(* IEC 61131-3 sources: SemaPLC/sema-plc-benchmark/spec2control-benchmark/data/st-baseline/steel-plant/pous/programs, 9 files *)

(* ---- main.st ---- *)
PROGRAM main
VAR
	Heartbeat : bool;
END_VAR

(* Entry point required by OpenPLC Editor v4. The process sections run as parallel program instances under task0; main only provides a scan heartbeat. *)
Heartbeat := NOT Heartbeat;

END_PROGRAM

(* ---- Section2.st ---- *)
PROGRAM Section2
VAR
	FT101_WildFlow_PV : real;
	FT102_FluxFlow_PV : real;
	TIT101_Temperature_PV : real;
	FFIC103_FluxFlow_SP : real;
	FT_101 : ANALOG_IN;
	FT_102 : ANALOG_IN;
	TIT_101 : ANALOG_IN;
	FFIC_103 : RATIO_CONTROL;
	FIC_102 : PID_BASIC;
	FV_102 : VALVE_ELECTRIC;
	LowFlow_OK_GT : bool;
	FFIC103_LowTempOrLowFlow_OR : bool;
	FFIC103_SensorFaults_OR : bool;
	FFIC103_RangeOrLowTempLowFlow_OR : bool;
	FFIC103_Inhibit_OR : bool;
END_VAR

FT_101(
    PV_Low := 50.0,
    Scaling_Slope := 62.5,
    Scaling_Offset := -250.0,
    Alarm_Enable := TRUE);
FT_102(
    Alarm_Enable := TRUE);
TIT_101(
    PV_Low := 800.0,
    Alarm_Enable := TRUE);
FFIC103_LowTempOrLowFlow_OR := FT_101.Low_Alarm OR TIT_101.Low_Alarm;
FFIC103_RangeOrLowTempLowFlow_OR := FT_101.High_Alarm OR FFIC103_LowTempOrLowFlow_OR;
FFIC103_SensorFaults_OR := FT_101.General_Fault OR FT_102.General_Fault;
FFIC103_Inhibit_OR := FFIC103_SensorFaults_OR OR FFIC103_RangeOrLowTempLowFlow_OR;
LowFlow_OK_GT := (FT_101.PV > 50.0);
FFIC_103(
    Auto := LowFlow_OK_GT,
    PrimaryPV := FT_101.PV,
    SecondaryPV := FT_102.PV,
    RatioSP := 0.4,
    MV_MIN := 200.0,
    MV_MAX := 300.0,
    Inhibit := FFIC103_Inhibit_OR);
FIC_102(
    AUTO := LowFlow_OK_GT,
    PV := FT_102.PV,
    SP := FFIC_103.SlaveSP);
FV_102(
    Control_Signal := FIC_102.XOUT,
    Inhibit := FFIC103_LowTempOrLowFlow_OR);

(* Outputs published to other sections / HMI. *)
FT101_WildFlow_PV := FT_101.PV;
FT102_FluxFlow_PV := FT_102.PV;
TIT101_Temperature_PV := TIT_101.PV;
FFIC103_FluxFlow_SP := FFIC_103.SlaveSP;

END_PROGRAM

(* ---- Section3.st ---- *)
PROGRAM Section3
VAR
	PT_201_VOTE_PV : real;
	TT_201_VOTE_PV : real;
	PT_201A : ANALOG_IN;
	PT_201B : ANALOG_IN;
	PT_201C : ANALOG_IN;
	TT_201A : ANALOG_IN;
	TT_201B : ANALOG_IN;
	TT_201C : ANALOG_IN;
	PT_201_VOTE : VOTING_ANALOG;
	TT_201_VOTE : VOTING_ANALOG;
	P_201 : MOTOR_ON_OFF;
	MO_201 : DIGITAL_IN;
	MO_202 : DIGITAL_IN;
	I_201 : BOOL_INPUT;
	I_202 : BOOL_INPUT;
	SI_201 : BOOL_INPUT;
	SI_202 : BOOL_INPUT;
	PT_GeneralFault : bool;
	MO201_Invert : bool;
	PT_SummaryPre : bool;
	PT_SummaryMasked : bool;
	TT_GeneralFault : bool;
	MO202_Invert : bool;
	TT_SummaryPre : bool;
	TT_SummaryMasked : bool;
	PressureInhibit : bool;
	TemperatureInhibit : bool;
	PumpInhibit : bool;
	PT_PressureHigh : bool;
	TT_TemperatureHigh : bool;
	PT_PressurePermissive : bool;
	TT_TemperaturePermissive : bool;
	StartPermissiveOK : bool;
	StartPermissiveNot : bool;
END_VAR

PT_201A(
    PV_High := 100.0,
    Alarm_Enable := TRUE);
PT_201B(
    PV_High := 100.0,
    Alarm_Enable := TRUE);
PT_201C(
    PV_High := 100.0,
    Alarm_Enable := TRUE);
TT_201A(
    Alarm_Enable := TRUE);
TT_201B(
    Alarm_Enable := TRUE);
TT_201C(
    Alarm_Enable := TRUE);
PT_PressureHigh := (PT_201_VOTE_PV > 100.0);
I_201(
    Bool_In := PT_PressureHigh,
    Alarm_OnTrue := TRUE,
    Latch_Enable := TRUE);
MO_201();
MO201_Invert := NOT MO_201.DI_Out;
PT_GeneralFault := PT_201A.General_Fault OR PT_201B.General_Fault OR PT_201C.General_Fault;
PT_SummaryPre := PT_GeneralFault OR PT_201_VOTE.Alarm_Voting_Error;
PT_SummaryMasked := PT_SummaryPre AND MO201_Invert;
SI_201(
    Bool_In := PT_SummaryMasked,
    Alarm_OnTrue := TRUE,
    Latch_Enable := TRUE);
PressureInhibit := I_201.Bool_Out OR SI_201.Bool_Out;
PT_201_VOTE(
    Input1 := PT_201A.PV,
    Input2 := PT_201B.PV,
    Input3 := PT_201C.PV,
    Deviation_Limit := 5.0,
    Voting_Scheme := '"2oo3"',
    EnableAlarm := TRUE,
    Inhibit := PressureInhibit);
TT_TemperatureHigh := (TT_201_VOTE_PV > 75.0);
I_202(
    Bool_In := TT_TemperatureHigh,
    Alarm_OnTrue := TRUE,
    Latch_Enable := TRUE);
MO_202();
MO202_Invert := NOT MO_202.DI_Out;
TT_GeneralFault := TT_201A.General_Fault OR TT_201B.General_Fault OR TT_201C.General_Fault;
TT_SummaryPre := TT_GeneralFault OR TT_201_VOTE.Alarm_Voting_Error;
TT_SummaryMasked := TT_SummaryPre AND MO202_Invert;
SI_202(
    Bool_In := TT_SummaryMasked,
    Alarm_OnTrue := TRUE,
    Latch_Enable := TRUE);
TemperatureInhibit := I_202.Bool_Out OR SI_202.Bool_Out;
TT_201_VOTE(
    Input1 := TT_201A.PV,
    Input2 := TT_201B.PV,
    Input3 := TT_201C.PV,
    Deviation_Limit := 5.0,
    Voting_Scheme := '"Median"',
    EnableAlarm := TRUE,
    Inhibit := TemperatureInhibit);
PT_PressurePermissive := (PT_201_VOTE_PV >= 21.0);
TT_TemperaturePermissive := (TT_201_VOTE_PV < 75.0);
StartPermissiveOK := PT_PressurePermissive AND TT_TemperaturePermissive;
StartPermissiveNot := NOT StartPermissiveOK;
PumpInhibit := TemperatureInhibit OR StartPermissiveNot;
P_201(
    Inhibit := PumpInhibit);

(* Outputs published to other sections / HMI. *)
PT_201_VOTE_PV := PT_201_VOTE.Voted_Output;
TT_201_VOTE_PV := TT_201_VOTE.Voted_Output;

END_PROGRAM

(* ---- Section4.st ---- *)
PROGRAM Section4
VAR
	FT_301_CoalFlow_PV : real;
	FT_302_AirFlow_PV : real;
	PT_301_Pressure_PV : real;
	TT_301_Temperature_PV : real;
	FIC_302_HotBlastAir_SP_FromRatio : real;
	Ratio_Bias : real;
	FT_301 : ANALOG_IN;
	PT_301 : ANALOG_IN;
	TT_301 : ANALOG_IN;
	FT_302 : ANALOG_IN;
	FFIC_303 : RATIO_CONTROL;
	FIC_302 : PID_BASIC;
	FV_302 : VALVE_ELECTRIC;
	FT301_Range_OR : bool;
	Shutdown_OR : bool;
	CombinedDisable_OR : bool;
	RatioInhibit_OR : bool;
	RatioAuto_NOT : bool;
	AirSP_Fallback_SEL : real;
	AirSP_Shutdown_SEL : real;
END_VAR

FT_301(
    PV_High := 5000.0,
    PV_Low := 100.0,
    Alarm_Enable := TRUE);
PT_301(
    Alarm_Enable := TRUE);
TT_301(
    Alarm_Enable := TRUE);
FT_302();
FT301_Range_OR := FT_301.High_Alarm OR FT_301.Low_Alarm;
Shutdown_OR := TT_301.Low_Alarm OR PT_301.High_Alarm;
CombinedDisable_OR := FT301_Range_OR OR Shutdown_OR;
RatioAuto_NOT := NOT CombinedDisable_OR;
RatioInhibit_OR := PT_301.High_Alarm OR TT_301.Low_Alarm OR FT_301.General_Fault OR PT_301.Low_Alarm;
FFIC_303(
    Auto := RatioAuto_NOT,
    PrimaryPV := FT_301.PV,
    SecondaryPV := FT_302.PV,
    RatioSP := 1.8,
    Bias := Ratio_Bias,
    TrimKp := 0.0,
    TrimTi := T#0s,
    MV_MIN := 200.0,
    MV_MAX := 9000.0,
    Inhibit := RatioInhibit_OR);
AirSP_Fallback_SEL := SEL(G := FT301_Range_OR, IN0 := FFIC_303.SlaveSP, IN1 := 500.0);
AirSP_Shutdown_SEL := SEL(G := Shutdown_OR, IN0 := AirSP_Fallback_SEL, IN1 := 0.0);
FIC_302(
    AUTO := TRUE,
    PV := FT_302.PV,
    SP := AirSP_Shutdown_SEL,
    MV_MIN := 0.0,
    MV_MAX := 100.0,
    X0 := 0.0,
    PV_High := 9000.0,
    PV_Low := 200.0,
    Inhibit := Shutdown_OR);
FV_302(
    Control_Signal := FIC_302.XOUT,
    Inhibit := Shutdown_OR);

(* Outputs published to other sections / HMI. *)
FT_301_CoalFlow_PV := FT_301.PV;
FT_302_AirFlow_PV := FT_302.PV;
PT_301_Pressure_PV := PT_301.PV;
TT_301_Temperature_PV := TT_301.PV;
FIC_302_HotBlastAir_SP_FromRatio := FFIC_303.SlaveSP;

END_PROGRAM

(* ---- Section5.st ---- *)
PROGRAM Section5
VAR
	TT_401_V_Temp_PV : real;
	PT_401_V_Pressure_PV : real;
	FT_401_Flow_PV : real;
	FT_401 : ANALOG_IN;
	PT_401A : ANALOG_IN;
	PT_401B : ANALOG_IN;
	PT_401C : ANALOG_IN;
	TT_401 : ANALOG_IN;
	TT_401A : ANALOG_IN;
	TT_401B : ANALOG_IN;
	TT_401C : ANALOG_IN;
	TT_401_V : VOTING_ANALOG;
	PT_401_V : VOTING_ANALOG;
	BOF_401_TempControl : PID_BASIC;
	BOF_402 : VALVE_ELECTRIC;
	I_401 : BOOL_INPUT;
	MA_401 : BOOL_INPUT;
	DA_401 : BOOL_INPUT;
	FA_401 : BOOL_INPUT;
	FlowPermissive_NOT : bool;
	PTA_HighAlarm_OK_NOT : bool;
	PTA_LowAlarm_OK_NOT : bool;
	PTB_HighAlarm_OK_NOT : bool;
	PTB_LowAlarm_OK_NOT : bool;
	PTC_HighAlarm_OK_NOT : bool;
	PTC_LowAlarm_OK_NOT : bool;
	PTA_WithinRange_AND : bool;
	PTB_WithinRange_AND : bool;
	PTC_WithinRange_AND : bool;
	PT_AB_Within_AND : bool;
	PT_AC_Within_AND : bool;
	PT_BC_Within_AND : bool;
	PT_2oo3_OK_OR1 : bool;
	PT_2oo3_OK_OR : bool;
	TempVoted_GT : bool;
	HealthySensors_GT : bool;
	TempPermit_AND : bool;
	AllPermissives_OK_AND1 : bool;
	AllPermissives_OK_AND : bool;
	PermissivesFail_NOT : bool;
	SensorFaults_OR1 : bool;
	SensorFaults_OR2 : bool;
	SensorFaults_OR3 : bool;
	SensorFaults_OR4 : bool;
	SensorFaults_OR5 : bool;
	SensorFaults_OR6 : bool;
	SensorFaults_OR7 : bool;
	Inhibit_OR1 : bool;
	Inhibit_OR : bool;
END_VAR

FT_401(
    Alarm_Enable := TRUE);
PT_401A(
    Alarm_Enable := TRUE);
PT_401B(
    Alarm_Enable := TRUE);
PT_401C(
    Alarm_Enable := TRUE);
TT_401(
    Alarm_Enable := TRUE);
TT_401A(
    Alarm_Enable := TRUE);
TT_401B(
    Alarm_Enable := TRUE);
TT_401C(
    Alarm_Enable := TRUE);
TT_401_V(
    Input1 := TT_401A.PV,
    Input2 := TT_401B.PV,
    Input3 := TT_401C.PV,
    Deviation_Limit := 0.05,
    Voting_Scheme := 'Median',
    EnableAlarm := TRUE);
PT_401_V(
    Input1 := PT_401A.PV,
    Input2 := PT_401B.PV,
    Input3 := PT_401C.PV,
    Voting_Scheme := '2oo3',
    EnableAlarm := TRUE);
BOF_401_TempControl(
    AUTO := TRUE,
    PV := TT_401_V.Voted_Output,
    SP := 1650.0,
    MV_MIN := 0.0,
    MV_MAX := 100.0,
    X0 := 0.0,
    KP := 1.0,
    TR := 60.0,
    TD := 0.0);
SensorFaults_OR1 := TT_401A.General_Fault OR TT_401B.General_Fault;
SensorFaults_OR2 := SensorFaults_OR1 OR TT_401C.General_Fault;
SensorFaults_OR3 := SensorFaults_OR2 OR TT_401.General_Fault;
SensorFaults_OR4 := SensorFaults_OR3 OR PT_401A.General_Fault;
SensorFaults_OR5 := SensorFaults_OR4 OR PT_401B.General_Fault;
SensorFaults_OR6 := SensorFaults_OR5 OR PT_401C.General_Fault;
SensorFaults_OR7 := SensorFaults_OR6 OR FT_401.General_Fault;
FA_401(
    Bool_In := SensorFaults_OR7);
DA_401(
    Bool_In := TT_401_V.Alarm_Voting_Error);
PTA_HighAlarm_OK_NOT := NOT PT_401A.High_Alarm;
PTA_LowAlarm_OK_NOT := NOT PT_401A.Low_Alarm;
PTA_WithinRange_AND := PTA_HighAlarm_OK_NOT AND PTA_LowAlarm_OK_NOT;
PTB_HighAlarm_OK_NOT := NOT PT_401B.High_Alarm;
PTB_LowAlarm_OK_NOT := NOT PT_401B.Low_Alarm;
PTB_WithinRange_AND := PTB_HighAlarm_OK_NOT AND PTB_LowAlarm_OK_NOT;
PT_AB_Within_AND := PTA_WithinRange_AND AND PTB_WithinRange_AND;
PTC_HighAlarm_OK_NOT := NOT PT_401C.High_Alarm;
PTC_LowAlarm_OK_NOT := NOT PT_401C.Low_Alarm;
PTC_WithinRange_AND := PTC_HighAlarm_OK_NOT AND PTC_LowAlarm_OK_NOT;
PT_AC_Within_AND := PTA_WithinRange_AND AND PTC_WithinRange_AND;
PT_2oo3_OK_OR1 := PT_AB_Within_AND OR PT_AC_Within_AND;
PT_BC_Within_AND := PTB_WithinRange_AND AND PTC_WithinRange_AND;
PT_2oo3_OK_OR := PT_2oo3_OK_OR1 OR PT_BC_Within_AND;
HealthySensors_GT := (TT_401_V.Healthy_Sensors_Count > 1);
TempVoted_GT := (TT_401_V.Voted_Output > 1450.0);
TempPermit_AND := TempVoted_GT AND HealthySensors_GT;
AllPermissives_OK_AND1 := TempPermit_AND AND PT_2oo3_OK_OR;
FlowPermissive_NOT := NOT FT_401.Low_Alarm;
AllPermissives_OK_AND := AllPermissives_OK_AND1 AND FlowPermissive_NOT;
PermissivesFail_NOT := NOT AllPermissives_OK_AND;
Inhibit_OR1 := PermissivesFail_NOT OR DA_401.Bool_Out;
Inhibit_OR := Inhibit_OR1 OR FA_401.Bool_Out;
I_401(
    Bool_In := Inhibit_OR);
BOF_402(
    Control_Signal := BOF_401_TempControl.XOUT,
    Manual_Mode := FALSE,
    Manual_Position := 0.0,
    Open_Limit := 100.0,
    Close_Limit := 0.0,
    Timeout := T#10s,
    Inhibit := I_401.Bool_Out);
MA_401();

(* Outputs published to other sections / HMI. *)
TT_401_V_Temp_PV := TT_401_V.Voted_Output;
PT_401_V_Pressure_PV := PT_401_V.Voted_Output;
FT_401_Flow_PV := FT_401.PV;

END_PROGRAM

(* ---- Section6.st ---- *)
PROGRAM Section6
VAR
	PT_501_Pressure_PV : real;
	TT_501_Temperature_PV : real;
	TT_501_MV : real;
	SM_501_EA_POS : real;
	SM_501_EA_CMD : real;
	PT_501 : ANALOG_IN;
	TT_501 : ANALOG_IN;
	SM_501 : VALVE_ELECTRIC;
	TT_501_CTRL : PID_BASIC;
	SM_501_LID_POS : DIGITAL_IN;
	HeatingEnableDelay_TON : TON;
	HeatingInhibit_OR : bool;
	LidNotClosed_NOT : bool;
	EAposLE10_LE : bool;
	HeatingEnableReq_NOT : bool;
	AutoMode_NOT : bool;
END_VAR

PT_501(
    Alarm_Enable := TRUE);
TT_501(
    PV_High := 1650.0,
    PV_Low := 1500.0,
    Scaling_Slope := 37.5,
    Scaling_Offset := 1050.0,
    Alarm_Enable := TRUE);
EAposLE10_LE := (SM_501.Feedback_Pos <= 10.0);
SM_501_LID_POS();
LidNotClosed_NOT := NOT SM_501_LID_POS.DI_Out;
HeatingInhibit_OR := LidNotClosed_NOT OR TT_501.High_Alarm OR PT_501.Low_Alarm OR TT_501.General_Fault OR SM_501.Alarm OR EAposLE10_LE;
HeatingEnableReq_NOT := NOT HeatingInhibit_OR;
HeatingEnableDelay_TON(
    IN := HeatingEnableReq_NOT,
    PT := T#10s);
AutoMode_NOT := NOT HeatingEnableDelay_TON.Q;
TT_501_CTRL(
    AUTO := HeatingEnableDelay_TON.Q,
    PV := TT_501.PV,
    SP := 1620.0,
    MV_MIN := 0.0,
    MV_MAX := 100.0,
    X0 := SM_501.Feedback_Pos,
    KP := 3.2,
    TR := 1.5,
    TD := 0.3,
    PV_High := 1650.0,
    PV_Low := 1500.0,
    Deviation_Limit := 2.0,
    Inhibit := HeatingInhibit_OR);
SM_501(
    Control_Signal := TT_501_CTRL.XOUT,
    Manual_Mode := AutoMode_NOT,
    Manual_Position := 0.0,
    Open_Limit := 100.0,
    Close_Limit := 0.0,
    Timeout := T#5s,
    Inhibit := HeatingInhibit_OR);

(* Outputs published to other sections / HMI. *)
PT_501_Pressure_PV := PT_501.PV;
TT_501_Temperature_PV := TT_501.PV;
TT_501_MV := TT_501_CTRL.XOUT;
SM_501_EA_POS := SM_501.Feedback_Pos;
SM_501_EA_CMD := SM_501.Valve_Position;

END_PROGRAM

(* ---- Section7.st ---- *)
PROGRAM Section7
VAR
	LIT101_MoldLevel_PV_mm : real;
	FT601_CoolingWaterFlow_PV_m3h : real;
	TT601_MoldTemp_PV_C : real;
	LIC101_ControllerOutput_Pct : real;
	LIT_101 : ANALOG_IN;
	FT_601 : ANALOG_IN;
	TT_601 : ANALOG_IN;
	LIC_101 : PID_BASIC;
	MV_101 : VALVE_ELECTRIC;
	ILK_FT_601_LOW : BOOL_INPUT;
	ILK_TT_601_HIGH : BOOL_INPUT;
	PERM_LIT_101_UNDER_250 : BOOL_INPUT;
	ILK_LIT_101_HIGH_HIGH_280 : BOOL_INPUT;
	ILK_LIT_101_FAULT : BOOL_INPUT;
	CC601_LoopTrips_OR : bool;
	MV101_Inhibit_OR : bool;
END_VAR

LIT_101(
    PV_High := 280.0,
    Scaling_Slope := 18.75,
    Scaling_Offset := -75.0,
    Alarm_Enable := TRUE);
FT_601(
    Alarm_Enable := TRUE);
TT_601(
    PV_High := 950.0,
    Alarm_Enable := TRUE);
ILK_FT_601_LOW(
    Bool_In := FT_601.Low_Alarm);
ILK_LIT_101_FAULT(
    Bool_In := LIT_101.General_Fault);
ILK_TT_601_HIGH(
    Bool_In := TT_601.High_Alarm);
CC601_LoopTrips_OR := ILK_FT_601_LOW.Bool_Out OR ILK_TT_601_HIGH.Bool_Out OR ILK_LIT_101_FAULT.Bool_Out;
ILK_LIT_101_HIGH_HIGH_280(
    Bool_In := LIT_101.High_Alarm);
PERM_LIT_101_UNDER_250(
    Bool_In := LIC_101.PV_High_Alarm);
MV101_Inhibit_OR := ILK_LIT_101_HIGH_HIGH_280.Bool_Out OR PERM_LIT_101_UNDER_250.Bool_Out OR CC601_LoopTrips_OR;
MV_101(
    Control_Signal := LIC_101.XOUT,
    Manual_Mode := FALSE,
    Open_Limit := 100.0,
    Close_Limit := 0.0,
    Inhibit := MV101_Inhibit_OR);
LIC_101(
    AUTO := TRUE,
    PV := LIT_101.PV,
    SP := 150.0,
    MV_MIN := 0.0,
    MV_MAX := 100.0,
    X0 := MV_101.Feedback_Pos,
    KP := -3.0,
    TR := 1.2,
    TD := 0.1,
    Deviation_Limit := 20.0,
    Inhibit := CC601_LoopTrips_OR);

(* Outputs published to other sections / HMI. *)
LIT101_MoldLevel_PV_mm := LIT_101.PV;
FT601_CoolingWaterFlow_PV_m3h := FT_601.PV;
TT601_MoldTemp_PV_C := TT_601.PV;
LIC101_ControllerOutput_Pct := LIC_101.XOUT;

END_PROGRAM

(* ---- Section8.st ---- *)
PROGRAM Section8
VAR
	FT701_FuelFlow_PV : real;
	FT702_AirFlow_PV : real;
	TT701_FurnaceTemp_PV : real;
	FLT701_FuelTankLevel_PV : real;
	FT702_SP_Ratio : real;
	FFIC701_ActiveRatio : real;
	FFIC701_RatioError : real;
	BLS701_BurnerStatus : bool;
	BLS701_BurnerStatus_DI : bool;
	ALM701_RatioAlarm : bool;
	ALM702_FT701Fault : bool;
	ALM703_FT702Fault : bool;
	ALM704_HighTemp : bool;
	FT_701 : ANALOG_IN;
	FT_702 : ANALOG_IN;
	TT_701 : ANALOG_IN;
	FLT_701 : ANALOG_IN;
	FFIC_701 : RATIO_CONTROL;
	FIC_702 : PID_BASIC;
	FV_702 : VALVE_ELECTRIC;
	BLS_701 : BOOL_INPUT;
	FuelGE200_GE : bool;
	BurnerOff_NOT : bool;
	TxFaults_OR : bool;
	FFICInhibit_OR1 : bool;
	FFICInhibit_OR2 : bool;
	FICInhibit_OR1 : bool;
	ValveInhibit_OR1 : bool;
	ValveInhibit_OR2 : bool;
	ValveInhibit_OR3 : bool;
	FFIC_Auto_AND1 : bool;
	FFIC_Auto_AND2 : bool;
	TempHigh_NOT : bool;
	RatioMinCalc_MULT : real;
	RatioMaxCalc_MULT : real;
	Ratio8xFuel_MULT : real;
	RatioLow_GT : bool;
	RatioHigh_GT : bool;
	RatioAlarm_OR : bool;
END_VAR

FT_701(
    Alarm_Enable := TRUE);
FT_702(
    Alarm_Enable := TRUE);
TT_701(
    PV_High := 1200.0,
    Alarm_Enable := TRUE);
FLT_701();
BLS_701(
    Bool_In := BLS701_BurnerStatus_DI,
    Alarm_OnTrue := FALSE,
    Alarm_OnFalse := TRUE,
    Latch_Enable := FALSE);
BurnerOff_NOT := NOT BLS_701.Bool_Out;
FFICInhibit_OR1 := BurnerOff_NOT OR FT_701.Low_Alarm;
TxFaults_OR := FT_701.General_Fault OR FT_702.General_Fault;
FFICInhibit_OR2 := FFICInhibit_OR1 OR TxFaults_OR;
FuelGE200_GE := (FT_701.PV >= 200.0);
FFIC_Auto_AND1 := FuelGE200_GE AND BLS_701.Bool_Out;
TempHigh_NOT := NOT TT_701.High_Alarm;
FFIC_Auto_AND2 := FFIC_Auto_AND1 AND TempHigh_NOT;
Ratio8xFuel_MULT := FT_701.PV * 8.0;
RatioMaxCalc_MULT := FT_701.PV * 12.0;
RatioMinCalc_MULT := FT_701.PV * 8.0;
FFIC_701(
    Auto := FFIC_Auto_AND2,
    PrimaryPV := FT_701.PV,
    SecondaryPV := FT_702.PV,
    RatioSP := 10.0,
    Bias := 0.0,
    MV_MIN := RatioMinCalc_MULT,
    MV_MAX := RatioMaxCalc_MULT,
    ManOut := Ratio8xFuel_MULT,
    Inhibit := FFICInhibit_OR2);
FICInhibit_OR1 := BurnerOff_NOT OR TxFaults_OR;
FIC_702(
    AUTO := TRUE,
    PV := FT_702.PV,
    SP := FFIC_701.SlaveSP,
    MV_MIN := 0.0,
    MV_MAX := 100.0,
    X0 := 0.0,
    KP := 1.5,
    TR := 10.0,
    TD := 0.5,
    Deviation_Limit := 5.0,
    Inhibit := FICInhibit_OR1);
ValveInhibit_OR1 := FT_701.Low_Alarm OR TT_701.Low_Alarm;
ValveInhibit_OR2 := ValveInhibit_OR1 OR TT_701.High_Alarm;
ValveInhibit_OR3 := ValveInhibit_OR2 OR TxFaults_OR;
FV_702(
    Control_Signal := FIC_702.XOUT,
    Manual_Mode := FALSE,
    Open_Limit := 100.0,
    Close_Limit := 0.0,
    Timeout := T#10s,
    Inhibit := ValveInhibit_OR3);
RatioLow_GT := (8.0 > FFIC_701.ActiveRatio);
RatioHigh_GT := (FFIC_701.ActiveRatio > 12.0);
RatioAlarm_OR := RatioLow_GT OR RatioHigh_GT;

(* Outputs published to other sections / HMI. *)
FT701_FuelFlow_PV := FT_701.PV;
FT702_AirFlow_PV := FT_702.PV;
TT701_FurnaceTemp_PV := TT_701.PV;
FLT701_FuelTankLevel_PV := FLT_701.PV;
FT702_SP_Ratio := FFIC_701.SlaveSP;
FFIC701_ActiveRatio := FFIC_701.ActiveRatio;
FFIC701_RatioError := FFIC_701.RatioErr;
BLS701_BurnerStatus := BLS_701.Bool_Out;
ALM702_FT701Fault := FT_701.General_Fault;
ALM703_FT702Fault := FT_702.General_Fault;
ALM704_HighTemp := TT_701.High_Alarm;
ALM701_RatioAlarm := RatioAlarm_OR;

END_PROGRAM

(* ---- Section9.st ---- *)
PROGRAM Section9
VAR
	FT801_Flow_PV : real;
	FT802_Flow_PV : real;
	PT801_Pressure_PV : real;
	FFIC801_AirFlow_SP : real;
	FFIC801_ActiveRatio : real;
	RatioHigh_Alarm : bool;
	RatioLow_Alarm : bool;
	AL_801 : ANALOG_IN;
	AL_802 : ANALOG_IN;
	AL_803 : ANALOG_IN;
	AL_804 : ANALOG_IN;
	FT_801 : ANALOG_IN;
	FT_802 : ANALOG_IN;
	PT_801 : ANALOG_IN;
	FFIC_801 : RATIO_CONTROL;
	FIC_802 : PID_BASIC;
	FV_802 : VALVE_ELECTRIC;
	RatioHighDelay_TON : TON;
	LowFlowEnable_GE : bool;
	PressureOutOfRange_OR : bool;
	FFIC801_Inhibits_OR : bool;
	FIC802_Faults_OR : bool;
	FV802_Inhibits_OR : bool;
	RatioHigh_GT : bool;
	RatioLow_LT : bool;
	NotFaults_NOT : bool;
	NotPressureLockout_NOT : bool;
	AutoEnable_AND : bool;
END_VAR

AL_801();
AL_802();
AL_803();
AL_804();
FT_801(
    Scaling_Slope := 312.5,
    Scaling_Offset := -1250.0,
    Alarm_Enable := TRUE);
FT_802(
    Scaling_Slope := 375.0,
    Scaling_Offset := -1500.0,
    Alarm_Enable := TRUE);
PT_801(
    Scaling_Slope := 0.125,
    Scaling_Offset := -0.5,
    Alarm_Enable := TRUE);
PressureOutOfRange_OR := PT_801.High_Alarm OR PT_801.Low_Alarm;
FFIC801_Inhibits_OR := PressureOutOfRange_OR OR FT_801.Low_Alarm OR FT_802.High_Alarm;
LowFlowEnable_GE := (FT_801.PV >= 100.0);
FFIC_801(
    Auto := LowFlowEnable_GE,
    PrimaryPV := FT_801.PV,
    SecondaryPV := FT_802.PV,
    RatioSP := 2.5,
    MV_MIN := 0.0,
    MV_MAX := 6000.0,
    Inhibit := FFIC801_Inhibits_OR);
FIC802_Faults_OR := FT_801.General_Fault OR PT_801.General_Fault;
NotFaults_NOT := NOT FIC802_Faults_OR;
NotPressureLockout_NOT := NOT PressureOutOfRange_OR;
AutoEnable_AND := LowFlowEnable_GE AND NotFaults_NOT AND NotPressureLockout_NOT;
FIC_802(
    AUTO := AutoEnable_AND,
    PV := FT_802.PV,
    SP := FFIC_801.SlaveSP,
    MV_MIN := 0.0,
    MV_MAX := 100.0,
    X0 := 50.0,
    Inhibit := FIC802_Faults_OR);
FV802_Inhibits_OR := PressureOutOfRange_OR OR FIC802_Faults_OR;
FV_802(
    Control_Signal := FIC_802.XOUT,
    Manual_Mode := PressureOutOfRange_OR,
    Manual_Position := 0.0,
    Open_Limit := 100.0,
    Close_Limit := 0.0,
    Inhibit := FV802_Inhibits_OR);
RatioHigh_GT := (FFIC_801.ActiveRatio > 3.0);
RatioHighDelay_TON(
    IN := RatioHigh_GT,
    PT := T#5s);
RatioLow_LT := (FFIC_801.ActiveRatio < 2.0);

(* Outputs published to other sections / HMI. *)
RatioHigh_Alarm := RatioHighDelay_TON.Q;
RatioLow_Alarm := RatioLow_LT;
FT801_Flow_PV := FT_801.PV;
FT802_Flow_PV := FT_802.PV;
PT801_Pressure_PV := PT_801.PV;
FFIC801_AirFlow_SP := FFIC_801.SlaveSP;
FFIC801_ActiveRatio := FFIC_801.ActiveRatio;

END_PROGRAM
